Fanuc KAREL source: kb00014.KL

PROGRAM KB00014
%STACKSIZE=65535
%PRIORITY=65535
%NOLOCKGROUP
VAR
P1 : FILE
RESULT : INTEGER
BEGIN
RESULT=BYTES_LEFT(P1)
END KB00014
